// IAG50cm#92: a stop during the HA stage of a park, on mock axes (IAG50cmTests README). Unlike the characterization suites this is
// a regression test of a defect: it FAILS until #92 is fixed. Every test owns a rig and runs over many PLC cycles (VAR_INST of the
// method, one Scan() per cycle). Failed checks are also noted in GVL_Diag.sFailures (printed by Run-Tests.ps1).
FUNCTION_BLOCK IagStopDuringPark_Tests EXTENDS TcUnit.FB_TestSuite
VAR
	fDecAtStop	: LREAL;		// Dec actual position when the stop was sent
END_VAR

Stop_Right_After_The_HA_Stage_Of_A_Park_Still_Stops_Dec();

// #92 (T18.4): the park moves HA home first, then commands the Dec move (MoveAxis -> fbAxis.MoveTo()). The NC reports InMotion a few
// cycles later (mock: SetStartScans), so for those scans both axes still report StandStill (bStopped). A stop in that window runs for one
// scan only: bStop is cleared at once (bStopped), the first scan of _StopTelescope only drops MoveAxis (CancelMove does not
// stop a move that was already started) and the axis stop (StopAxis) is never sent. The Dec move to home runs to the end.
// Expected: Dec is sent a stop and stays where it was. (A stop before the Dec command works: TCS_command passes stop and Dec never starts.)
// CI trace of the defect (TCS_command, bStop, bStopped, bPark, Dec MoveAxis, Dec InMotion): park 2, 0,1,1,1,0 -> stop 5, 0,1,0,0,0 -> no_command 0, 0,1,0,0,0
// -> then Dec InMotion for the rest of its 60 scan move with bStopped FALSE and no stop sent.
METHOD PRIVATE Stop_Right_After_The_HA_Stage_Of_A_Park_Still_Stops_Dec
VAR_INST
	rig			: FB_IagRig;
	nStep		: INT;
	nCycles		: UINT;
	bHaMoved	: BOOL;
	bSawStop	: BOOL;
	sTest		: STRING(80);
END_VAR
TEST('Stop_Right_After_The_HA_Stage_Of_A_Park_Still_Stops_Dec');
sTest := 'Stop_Right_After_The_HA_Stage_Of_A_Park_Still_Stops_Dec: ';
IF nStep >= 90 THEN
	RETURN;
END_IF
rig.Scan();
nCycles := nCycles + 1;
CASE nStep OF
0:	// wait for the clock, then power on
	IF rig.ClockValid THEN
		rig.fbTel.Init();
		rig.SetStartScans(nScans := 3);
		nStep := 10;
		nCycles := 0;
	ELSIF nCycles > 2000 THEN
		AssertTrue(Condition := FALSE, Message := 'the astronomical clock never became valid');
		F_Note(bFailed := TRUE, sText := CONCAT(sTest, 'the astronomical clock never became valid'));
		nStep := 99;
		TEST_FINISHED();
	END_IF
10:	// ready: slew away from home to a point with an hour angle, so that the park moves HA first
	IF rig.Online THEN
		rig.fbTel.Slew(fAzimuth := 120.0, fAltitude := 40.0);
		nStep := 20;
		nCycles := 0;
	ELSIF nCycles > 1500 THEN
		AssertTrue(Condition := FALSE, Message := 'the mock telescope did not reach READY_STATE 1.0');
		F_Note(bFailed := TRUE, sText := CONCAT(sTest, 'the mock telescope did not reach READY_STATE 1.0'));
		nStep := 99;
		TEST_FINISHED();
	END_IF
20:	// the slew has finished and the mount stands still: park
	IF nCycles > 10 AND NOT rig.fbTel.bSlewActive AND rig.fbTel.bStopped AND rig.fbTel.TCS_command <> E_TCSCommand.slew THEN
		rig.fbTel.Park();
		nStep := 30;
		nCycles := 0;
	ELSIF nCycles > 600 THEN
		AssertTrue(Condition := FALSE, Message := 'the slew did not finish');
		F_Note(bFailed := TRUE, sText := CONCAT(sTest, 'the slew did not finish'));
		nStep := 99;
		TEST_FINISHED();
	END_IF
30:	// wait until HA has been moved by the park and the Dec move is commanded but the axis does not report InMotion yet: stop now
	IF rig.fbHa.MoveAxis THEN
		bHaMoved := TRUE;
	END_IF
	IF bHaMoved AND rig.fbDec.MoveAxis AND NOT rig.fbDec.fbAxis.InMotion AND rig.fbTel.bParkActive THEN
		fDecAtStop := rig.fbDec.fActualPosition;
		rig.fbTel.Stop();
		nStep := 40;
		nCycles := 0;
	ELSIF NOT rig.fbTel.bParkActive AND nCycles > 5 THEN
		AssertTrue(Condition := FALSE, Message := 'the park ended before the HA stage could be observed');
		F_Note(bFailed := TRUE, sText := CONCAT(sTest, 'the park ended before the HA stage could be observed'));
		nStep := 99;
		TEST_FINISHED();
	ELSIF nCycles > 600 THEN
		AssertTrue(Condition := FALSE, Message := 'the park never finished its HA stage');
		F_Note(bFailed := TRUE, sText := CONCAT(sTest, 'the park never finished its HA stage'));
		nStep := 99;
		TEST_FINISHED();
	END_IF
40:	// the mock Dec move takes 60 scans: look when it would have ended
	IF rig.fbTel.TCS_command = E_TCSCommand.stop THEN
		bSawStop := TRUE;
	END_IF
	IF nCycles >= 100 THEN
		AssertTrue(Condition := bSawStop, Message := 'the stop command ran (TCS_command passed stop)');
		F_Note(bFailed := NOT (bSawStop), sText := CONCAT(sTest, 'the stop command ran (TCS_command passed stop)'));
		AssertFalse(Condition := rig.fbTel.bParkActive, Message := 'the park is cancelled');
		F_Note(bFailed := (rig.fbTel.bParkActive), sText := CONCAT(sTest, 'the park is cancelled'));
		AssertTrue(Condition := rig.fbDec.nStopEdges >= 1, Message := 'Dec was sent an axis stop (the Dec move had started)');
		F_Note(bFailed := NOT (rig.fbDec.nStopEdges >= 1), sText := CONCAT(sTest, 'Dec was sent an axis stop (the Dec move had started)'));
		AssertTrue(Condition := rig.fbDec.fActualPosition = fDecAtStop, Message := 'Dec did not move to home after the stop');
		F_Note(bFailed := NOT (rig.fbDec.fActualPosition = fDecAtStop), sText := CONCAT(sTest, 'Dec did not move to home after the stop'));
		nStep := 99;
		TEST_FINISHED();
	END_IF
END_CASE
END_METHOD

END_FUNCTION_BLOCK

(* stored: Version 1.1.0.1, ProductVersion 3.1.4024.15
   POU IagStopDuringPark_Tests: Id {a12c82c6-ea41-4faa-936c-0cf6bcd4a223}, SpecialFunc None
   Method Stop_Right_After_The_HA_Stage_Of_A_Park_Still_Stops_Dec: Id {19d29f7c-7cb6-48a5-8673-fd458202fb79} *)
